Staubli VAL3: getPointPara.pgx

public program getPointPara(string x_sKey, num x_nIndex, num& x_nMoveType, num& x_nParaSpeed, num& x_nParaAccel, num& x_nParaBlend, num x_nParaPercent, string& x_sComment, bool& x_bSafePoint, string& x_sBlend, num& x_nValue[], string& x_sTRSF[])
  local num l_nMoveType
begin
  x_nMoveType=trajTemp:tTrajItem[x_sKey].pPointItem[x_nIndex].pParaItem.nMoveType
  x_nParaSpeed=trajTemp:tTrajItem[x_sKey].pPointItem[x_nIndex].pParaItem.mMdesc.vel
  x_nParaAccel=trajTemp:tTrajItem[x_sKey].pPointItem[x_nIndex].pParaItem.mMdesc.accel
  x_nParaBlend=trajTemp:tTrajItem[x_sKey].pPointItem[x_nIndex].pParaItem.mMdesc.leave
  x_nParaPercent=trajTemp:tTrajItem[x_sKey].pPointItem[x_nIndex].pParaItem.nPercentage
  x_sComment=trajTemp:tTrajItem[x_sKey].pPointItem[x_nIndex].sID
  //  x_bBlendJoint=(trajTemp:tTrajItem[x_sKey].pPointItem[x_nIndex].pParaItem.mMdesc.blend==joint)
  //  x_bBlendOFF=(trajTemp:tTrajItem[x_sKey].pPointItem[x_nIndex].pParaItem.mMdesc.blend==off)
  switch x_nMoveType
    case 1

      x_nValue[0]=trajTemp:tTrajItem[x_sKey].pPointItem[x_nIndex].jJointRx.j1
      x_nValue[1]=trajTemp:tTrajItem[x_sKey].pPointItem[x_nIndex].jJointRx.j2
      x_nValue[2]=trajTemp:tTrajItem[x_sKey].pPointItem[x_nIndex].jJointRx.j3
      x_nValue[3]=trajTemp:tTrajItem[x_sKey].pPointItem[x_nIndex].jJointRx.j4
      x_nValue[4]=trajTemp:tTrajItem[x_sKey].pPointItem[x_nIndex].jJointRx.j5
      x_nValue[5]=trajTemp:tTrajItem[x_sKey].pPointItem[x_nIndex].jJointRx.j6

      x_sTRSF[0]="J1:"
      x_sTRSF[1]="J2:"
      x_sTRSF[2]="J3:"
      x_sTRSF[3]="J4:"
      x_sTRSF[4]="J5:"
      x_sTRSF[5]="J6:"

    break
    case 0
      x_nValue[0]=trajTemp:tTrajItem[x_sKey].pPointItem[x_nIndex].pPointRx.trsf.x
      x_nValue[1]=trajTemp:tTrajItem[x_sKey].pPointItem[x_nIndex].pPointRx.trsf.y
      x_nValue[2]=trajTemp:tTrajItem[x_sKey].pPointItem[x_nIndex].pPointRx.trsf.z
      x_nValue[3]=trajTemp:tTrajItem[x_sKey].pPointItem[x_nIndex].pPointRx.trsf.rx
      x_nValue[4]=trajTemp:tTrajItem[x_sKey].pPointItem[x_nIndex].pPointRx.trsf.ry
      x_nValue[5]=trajTemp:tTrajItem[x_sKey].pPointItem[x_nIndex].pPointRx.trsf.rz

      x_sTRSF[0]="X:"
      x_sTRSF[1]="Y:"
      x_sTRSF[2]="Z:"
      x_sTRSF[3]="RX:"
      x_sTRSF[4]="RY:"
      x_sTRSF[5]="RZ:"
    break
    case 2
      x_nValue[0]=trajTemp:tTrajItem[x_sKey].pPointItem[x_nIndex].pPointRx.trsf.x
      x_nValue[1]=trajTemp:tTrajItem[x_sKey].pPointItem[x_nIndex].pPointRx.trsf.y
      x_nValue[2]=trajTemp:tTrajItem[x_sKey].pPointItem[x_nIndex].pPointRx.trsf.z
      x_nValue[3]=trajTemp:tTrajItem[x_sKey].pPointItem[x_nIndex].pPointRx.trsf.rx
      x_nValue[4]=trajTemp:tTrajItem[x_sKey].pPointItem[x_nIndex].pPointRx.trsf.ry
      x_nValue[5]=trajTemp:tTrajItem[x_sKey].pPointItem[x_nIndex].pPointRx.trsf.rz
      x_nValue[6]= trajTemp:tTrajItem[x_sKey].pPointItem[x_nIndex].pInter.trsf.x
      x_nValue[7]=trajTemp:tTrajItem[x_sKey].pPointItem[x_nIndex].pInter.trsf.y
      x_nValue[8]=trajTemp:tTrajItem[x_sKey].pPointItem[x_nIndex].pInter.trsf.z
      x_nValue[9]=trajTemp:tTrajItem[x_sKey].pPointItem[x_nIndex].pInter.trsf.rx
      x_nValue[10]=trajTemp:tTrajItem[x_sKey].pPointItem[x_nIndex].pInter.trsf.ry
      x_nValue[11]= trajTemp:tTrajItem[x_sKey].pPointItem[x_nIndex].pInter.trsf.rz
      x_sTRSF[0]="X:"
      x_sTRSF[1]="Y:"
      x_sTRSF[2]="Z:"
      x_sTRSF[3]="RX:"
      x_sTRSF[4]="RY:"
      x_sTRSF[5]="RZ:"
      x_sTRSF[6]="2X:"
      x_sTRSF[7]="2Y:"
      x_sTRSF[8]="2Z:"
      x_sTRSF[9]="2RX:"
      x_sTRSF[10]="2RY:"
      x_sTRSF[11]="2RZ:"

    break
  endSwitch
  //blend
  if trajTemp:tTrajItem[x_sKey].pPointItem[x_nIndex].pParaItem.mMdesc.blend==off
    x_sBlend="OFF"
  elseIf trajTemp:tTrajItem[x_sKey].pPointItem[x_nIndex].pParaItem.mMdesc.blend==joint
    x_sBlend="关节"
  elseIf trajTemp:tTrajItem[x_sKey].pPointItem[x_nIndex].pParaItem.mMdesc.blend==Cartesian
    x_sBlend="笛卡尔"
  endIf
  x_bSafePoint = (trajTemp:tTrajItem[x_sKey].pPointItem.pParaItem.bSafePoint==true)
end
